Fanuc KAREL source: ka00133.KL

PROGRAM KA00133
%STACKSIZE=65535
%PRIORITY=65535
%NOLOCKGROUP
VAR
SRC : ARRAY[2] OF SHORT
DST : INTEGER
BEGIN
SRC[1]=2
DST=SRC[1]
END KA00133
